{attribute 'linkalways'}
{attribute 'no_explicit_call' := 'This FB is a CLASS and must be accessed using methods or properties'}
{attribute 'enable_dynamic_creation'}
FUNCTION_BLOCK Node_F_VN_InnerCircle EXTENDS VisionNode
VAR
    ipSrcImage : _ITcVnImage;
    fRadius : _LREAL(0.0);
    aCenter : _TcVnPoint2_REAL;
    hrPrev : _HRESULT(S_OK);
    hresult : _HRESULT(S_OK);
END_VAR

METHOD PUBLIC Clone : I_Node
VAR
    pNode : POINTER TO Node_F_VN_InnerCircle;
END_VAR
pNode := __NEW(Node_F_VN_InnerCircle);
Clone := pNode^;
END_METHOD

METHOD FB_init : BOOL
VAR_INPUT
    bInitRetains : BOOL;
    bInCopyCode : BOOL;
END_VAR
AddInput('ipSrcImage', ipSrcImage);
AddInput('hrPrev', hrPrev);
AddOutput('fRadius', fRadius);
AddOutput('aCenter', aCenter);
AddOutput('hresult', hresult);
END_METHOD

METHOD PROTECTED OnExecute
hresult.Value := F_VN_InnerCircle(
    ipSrcImage := ipSrcImage.Value,
    fRadius := fRadius.Value,
    aCenter := aCenter.Value,
    hrPrev := hrPrev.Value);
END_METHOD

METHOD PUBLIC PreExecutionCheck
VAR_INPUT
    Check : I_PreExecutionChecks;
END_VAR
Check.IsTrue(ipSrcImage.IsValid, 'ipSrcImage must contain an image');
Check.IsTrue(ipSrcImage.HasChannelCount(1), 'ipSrcImage must have 1 channel');
Check.IsTrue(ipSrcImage.IsElementType(ETcVnElementType.TCVN_ET_USINT), 'ipSrcImage must contain USINT elements');
END_METHOD

END_FUNCTION_BLOCK

(* stored: Version 1.1.0.1, ProductVersion 3.1.4026.19
   POU Node_F_VN_InnerCircle: Id {469575f2-633a-4e7d-a6c1-8010eb5168df}, SpecialFunc None
   Folder Constructor: Id {64ad9d86-fa54-42d5-ae81-d072d1dcc004}
   Method Clone: Id {e8549939-342e-45d3-85a0-cb6a22c4d0af}
   Method FB_init: Id {bdabecd7-0a71-453a-ad12-16705f1f65d3}
   Method OnExecute: Id {56c0e4dd-3a49-4cde-be69-ff73078a0c51}
   Method PreExecutionCheck: Id {af200c86-070e-43f9-800e-0c8c8705c3b4} *)
